// TIA Portal V20 export
Screen "190RB02_V23"  1276x673
  ScreenItem "Line_Header_X0_Y64" at 0,64 size 1276x0  Type=HmiLine
  ScreenItem "permanentareaborderrectangle" at 0,0 size 0x0  Type=HmiRectangle
  ScreenItem "Button_Back" at 2,2 size 90x60  Type=HmiButton
  ScreenItem "Title_ScreenOverview_X390_Y2_2" at 392,5 size 510x57  Type=HmiTextBox
  ScreenItem "Fusszeile_Button_ManualOPMode1_4" at 1181,2 size 90x60  Type=HmiButton
  ScreenItem "Title_ScreenOverview_X390_Y2_1" at 1130,78 size 139x57  Type=HmiTextBox
  ScreenItem "Title_ScreenOverview_X390_Y2_3" at 1130,144 size 139x57  Type=HmiTextBox
  ScreenItem "Title_ScreenOverview_X390_Y2_4" at 1130,144 size 139x57  Type=HmiTextBox
  ScreenItem "Graphic view_2" at 215,99 size 741x526  Type=HmiGraphicView
  ScreenItem "Line_4" at 603,164 size 56x114  Type=HmiLine
  ScreenItem "文本域_11" at 623,75 size 134x40  Type=HmiTextBox
  ScreenItem "Line_10" at 858,213 size 105x69  Type=HmiLine
  ScreenItem "文本域_1" at 990,242 size 134x40  Type=HmiTextBox
  ScreenItem "Line_1" at 912,300 size 81x29  Type=HmiLine
  ScreenItem "文本域_2" at 990,334 size 134x40  Type=HmiTextBox
  ScreenItem "Line_2" at 920,389 size 73x3  Type=HmiLine
  ScreenItem "文本域_3" at 971,431 size 134x40  Type=HmiTextBox
  ScreenItem "Line_3" at 807,368 size 154x97  Type=HmiLine
  ScreenItem "文本域_4" at 874,515 size 134x40  Type=HmiTextBox
  ScreenItem "Line_5" at 691,377 size 172x149  Type=HmiLine
  ScreenItem "文本域_5" at 640,526 size 134x40  Type=HmiTextBox
  ScreenItem "Line_6" at 612,444 size 73x74  Type=HmiLine
  ScreenItem "文本域_6" at 258,526 size 134x40  Type=HmiTextBox
  ScreenItem "Line_7" at 327,373 size 186x145  Type=HmiLine
  ScreenItem "Line_8" at 466,452 size 23x91  Type=HmiLine
  ScreenItem "文本域_7" at 398,552 size 134x40  Type=HmiTextBox
  ScreenItem "Line_9" at 148,411 size 130x67  Type=HmiLine
  ScreenItem "文本域_8" at 75,482 size 134x40  Type=HmiTextBox
  ScreenItem "文本域_9" at 28,377 size 134x40  Type=HmiTextBox
  ScreenItem "Line_11" at 164,361 size 113x52  Type=HmiLine
  ScreenItem "文本域_10" at 14,268 size 134x40  Type=HmiTextBox
  ScreenItem "Line_12" at 150,304 size 124x7  Type=HmiLine
  ScreenItem "Line_13" at 218,149 size 121x209  Type=HmiLine
  ScreenItem "文本域_13" at 245,99 size 134x40  Type=HmiTextBox
  ScreenItem "Line_14" at 326,196 size 96x148  Type=HmiLine
  ScreenItem "Line_15" at 463,182 size 36x83  Type=HmiLine
  ScreenItem "文本域_14" at 399,92 size 134x40  Type=HmiTextBox
  ScreenItem "Fusszeile_Button_ManualOPMode1_1" at 1088,2 size 90x60  Type=HmiButton
  ScreenItem "Title_ScreenOverview_X390_Y2_44" at 285,139 size 52x19  Type=HmiTextBox
  ScreenItem "Title_ScreenOverview_X390_Y2_45" at 285,159 size 25x21  Type=HmiTextBox
  ScreenItem "Title_ScreenOverview_X390_Y2_46" at 312,159 size 25x21  Type=HmiTextBox
  ScreenItem "Title_ScreenOverview_X390_Y2_5" at 437,132 size 52x19  Type=HmiTextBox
  ScreenItem "Title_ScreenOverview_X390_Y2_6" at 437,152 size 25x21  Type=HmiTextBox
  ScreenItem "Title_ScreenOverview_X390_Y2_7" at 464,152 size 25x21  Type=HmiTextBox
  ScreenItem "Title_ScreenOverview_X390_Y2_8" at 1061,302 size 25x21  Type=HmiTextBox
  ScreenItem "Title_ScreenOverview_X390_Y2_9" at 1034,282 size 52x19  Type=HmiTextBox
  ScreenItem "Title_ScreenOverview_X390_Y2_10" at 1034,302 size 25x21  Type=HmiTextBox
  ScreenItem "Title_ScreenOverview_X390_Y2_11" at 696,135 size 25x21  Type=HmiTextBox
  ScreenItem "Title_ScreenOverview_X390_Y2_12" at 669,115 size 52x19  Type=HmiTextBox
  ScreenItem "Title_ScreenOverview_X390_Y2_13" at 669,135 size 25x21  Type=HmiTextBox
  ScreenItem "Title_ScreenOverview_X390_Y2_14" at 1033,374 size 52x19  Type=HmiTextBox
  ScreenItem "Title_ScreenOverview_X390_Y2_15" at 1033,394 size 25x21  Type=HmiTextBox
  ScreenItem "Title_ScreenOverview_X390_Y2_16" at 1060,394 size 25x21  Type=HmiTextBox
  ScreenItem "Title_ScreenOverview_X390_Y2_17" at 1015,471 size 52x19  Type=HmiTextBox
  ScreenItem "Title_ScreenOverview_X390_Y2_18" at 1015,491 size 25x21  Type=HmiTextBox
  ScreenItem "Title_ScreenOverview_X390_Y2_19" at 1042,491 size 25x21  Type=HmiTextBox
  ScreenItem "Title_ScreenOverview_X390_Y2_20" at 922,556 size 52x19  Type=HmiTextBox
  ScreenItem "Title_ScreenOverview_X390_Y2_21" at 922,576 size 25x21  Type=HmiTextBox
  ScreenItem "Title_ScreenOverview_X390_Y2_22" at 949,576 size 25x21  Type=HmiTextBox
  ScreenItem "Title_ScreenOverview_X390_Y2_23" at 688,566 size 52x19  Type=HmiTextBox
  ScreenItem "Title_ScreenOverview_X390_Y2_24" at 688,586 size 25x21  Type=HmiTextBox
  ScreenItem "Title_ScreenOverview_X390_Y2_25" at 715,586 size 25x21  Type=HmiTextBox
  ScreenItem "Title_ScreenOverview_X390_Y2_26" at 432,613 size 25x21  Type=HmiTextBox
  ScreenItem "Title_ScreenOverview_X390_Y2_27" at 459,613 size 25x21  Type=HmiTextBox
  ScreenItem "Title_ScreenOverview_X390_Y2_28" at 432,593 size 52x19  Type=HmiTextBox
  ScreenItem "Title_ScreenOverview_X390_Y2_29" at 297,566 size 52x19  Type=HmiTextBox
  ScreenItem "Title_ScreenOverview_X390_Y2_30" at 297,586 size 25x21  Type=HmiTextBox
  ScreenItem "Title_ScreenOverview_X390_Y2_31" at 324,586 size 25x21  Type=HmiTextBox
  ScreenItem "Title_ScreenOverview_X390_Y2_32" at 115,526 size 52x19  Type=HmiTextBox
  ScreenItem "Title_ScreenOverview_X390_Y2_33" at 115,546 size 25x21  Type=HmiTextBox
  ScreenItem "Title_ScreenOverview_X390_Y2_34" at 142,546 size 25x21  Type=HmiTextBox
  ScreenItem "Title_ScreenOverview_X390_Y2_35" at 72,423 size 52x19  Type=HmiTextBox
  ScreenItem "Title_ScreenOverview_X390_Y2_36" at 72,443 size 25x21  Type=HmiTextBox
  ScreenItem "Title_ScreenOverview_X390_Y2_37" at 99,443 size 25x21  Type=HmiTextBox
  ScreenItem "Title_ScreenOverview_X390_Y2_38" at 83,333 size 25x21  Type=HmiTextBox
  ScreenItem "Title_ScreenOverview_X390_Y2_39" at 56,313 size 52x19  Type=HmiTextBox
  ScreenItem "Title_ScreenOverview_X390_Y2_40" at 56,333 size 25x21  Type=HmiTextBox
  ScreenItem "Rectangle_1" at 0,0 size 152x48  Type=HmiRectangle
  ScreenItem "文本域_15" at 2,1 size 122x45  Type=HmiTextBox
  ScreenItem "圆_1" at 0,0 size 100x30  Type=HmiCircle
  ScreenItem "圆_2" at 0,0 size 100x30  Type=HmiCircle
  ScreenItem "Rectangle_2" at 0,0 size 152x48  Type=HmiRectangle
  ScreenItem "文本域_16" at 2,1 size 122x45  Type=HmiTextBox
  ScreenItem "圆_3" at 0,0 size 100x30  Type=HmiCircle
  ScreenItem "圆_4" at 0,0 size 100x30  Type=HmiCircle
